(* IEC 61131-3 sources: SemantiST/compiler/intake/normalize/probes/scl-data-block, 2 files *)

(* ---- rewritten.st ---- *)
VAR_GLOBAL
SETTINGS :
{ S7_Optimized_Access := 'FALSE' }
(* VERSION : 0.1 *)
(* NON_RETAIN *)
   STRUCT
      LIMIT_HI : INT := 20;
      COUNT : INT;
   END_STRUCT;
END_VAR
   (* LIMIT_HI := 20; *)
(* END_DATA_BLOCK *)

FUNCTION main : DINT
SETTINGS.COUNT := 2;
printf('%d$N', SETTINGS.LIMIT_HI + SETTINGS.COUNT);
main := 0;
END_FUNCTION

(* ---- original.st ---- *)
DATA_BLOCK SETTINGS
{ S7_Optimized_Access := 'FALSE' }
VERSION : 0.1
NON_RETAIN
   STRUCT
      LIMIT_HI : INT := 10;
      COUNT : INT;
   END_STRUCT;
BEGIN
   LIMIT_HI := 20;
END_DATA_BLOCK

FUNCTION main : DINT
SETTINGS.COUNT := 2;
printf('%d$N', SETTINGS.LIMIT_HI + SETTINGS.COUNT);
main := 0;
END_FUNCTION
